ABB RAPID module: PgProg.prg

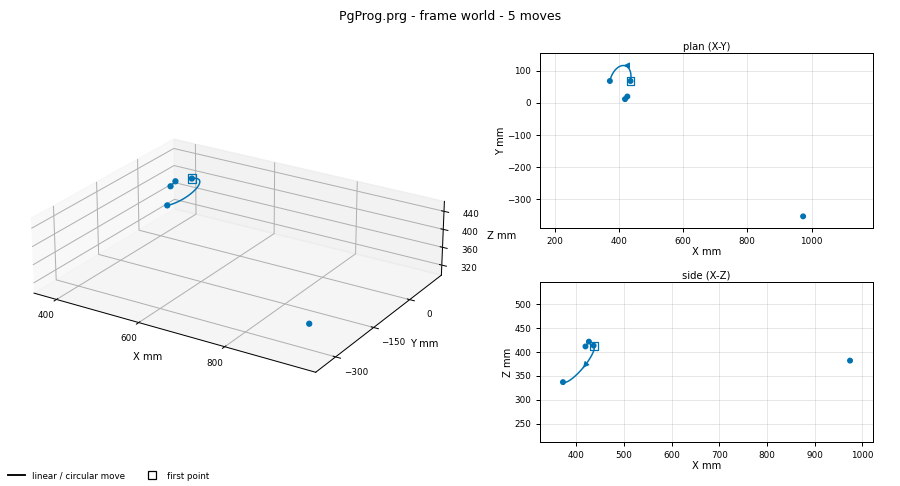
[picture p0: tool path of PgProg.prg in frame world, 5 of 9 moves have a stored position in this frame; points joined in program order, loops and branches not executed]
%%%
  VERSION:1
  LANGUAGE:ENGLISH
%%%
MODULE MOD_PgProg

    ! -------------------------------
    ! Define customized variables here
    ! ...

	! Tool variables:
	PERS tooldata ToolPg := [TRUE,[[10.000,20.000,150.000],[0.99144486,0.13052619,0.00000000,0.00000001]],[1,[0,0,20],[1,0,0,0],0,0,0.005]];
	PERS tooldata Tool2 := [TRUE,[[0.000,0.000,200.000],[1.00000000,0.00000000,0.00000000,0.00000000]],[1,[0,0,20],[1,0,0,0],0,0,0.005]];

	! Reference variables:
	PERS wobjdata FramePg := [FALSE, TRUE, "", [[1234.570,-98.765,50.500],[0.96592583,0.00000000,0.00000000,0.25881905]],[[0,0,0],[1,0,0,0]]];

	PROC Main()
		ConfJ \On;
		ConfL \Off;
		! Program generated by RoboDK v6.0.7 for ABB IRB 120-3/0.6 on XX/XX/XXXX 18:00:00
		! Using nominal kinematics.
		MoveAbsJ [[0.000000,-10.000000,20.000000,0.000000,30.000000,0.000000],[9E+09,9E+09,9E+09,9E+09,9E+09,9E+09]],[250.00,500,5000,1000],z5,ToolPg \WObj:=FramePg;
		MoveL [[-607.850,543.849,363.215],[0.37410804,0.28584607,0.85365954,-0.22271191],[0,0,0,0],[9E+09,9E+09,9E+09,9E+09,9E+09,9E+09]],[250.00,500,5000,1000],z5,ToolPg \WObj:=FramePg;
		MoveC [[-602.951,596.788,316.595],[0.37410804,0.28584607,0.85365954,-0.22271191],[0,0,0,0],[9E+09,9E+09,9E+09,9E+09,9E+09,9E+09]],[[-663.517,575.988,286.611],[0.37410804,0.28584607,0.85365954,-0.22271191],[0,0,0,0],[9E+09,9E+09,9E+09,9E+09,9E+09,9E+09]],[250.00,500,5000,1000],z5,ToolPg \WObj:=FramePg;
		MoveAbsJ [[20.000000,-10.000000,20.000000,0.000000,30.000000,0.000000],[9E+09,9E+09,9E+09,9E+09,9E+09,9E+09]],[250.00,500,5000,1000],z5,ToolPg \WObj:=FramePg;
		MoveL [[-650.861,503.437,361.399],[0.37410804,0.28584607,0.85365954,-0.22271191],[0,0,0,0],[9E+09,9E+09,9E+09,9E+09,9E+09,9E+09]],v100,z5,ToolPg \WObj:=FramePg;
		MoveL [[-640.584,506.980,371.534],[0.37410804,0.28584607,0.85365954,-0.22271191],[0,0,0,0],[9E+09,9E+09,9E+09,9E+09,9E+09,9E+09]],v100,z0,ToolPg \WObj:=FramePg;
		WaitTime 0.500;
		STOP;
		TPWrite "Hello from postgen";
		! a comment
		SubProgram;
		CustomCode(42)
		ThreadProg
		SetDO D_OUT_1, 1;
		SetDO Valve, 0;
		SetAO A_OUT_3, 2.5;
		WaitDI D_IN_2, 1;
		WaitDI D_IN_4, 0, \MaxTime:=1.5;
		MoveAbsJ [[0.000000,-10.000000,20.000000,0.000000,30.000000,0.000000],[9E+09,9E+09,9E+09,9E+09,9E+09,9E+09]],v100,z0,Tool2 \WObj:=FramePg;
		MoveAbsJ [[10.000000,-5.000000,25.000000,5.000000,35.000000,5.000000],[9E+09,9E+09,9E+09,9E+09,9E+09,9E+09]],v100,z0,Tool2 \WObj:=FramePg;
		MoveL [[-353.026,-90.135,331.702],[0.34432926,0.04805561,0.93307257,-0.09221494],[-1,0,-1,0],[9E+09,9E+09,9E+09,9E+09,9E+09,9E+09]],v100,z0,Tool2 \WObj:=FramePg;
	ENDPROC

ENDMODULE
